(* PLC project conveyor_station.project, CODESYS CODESYS V3.5 SP22 Patch 4 *)
(* stored: creationDateTime 2026-11-23T00:04:54.4201515, modificationDateTime 2026-11-23T00:02:17.3371292 *)

PROGRAM PLC_PRG
  VAR
    START_BTN : BOOL;  (* physical NO button *)
    STOP_BTN : BOOL := TRUE;  (* physical NC button (TRUE = not pressed) *)
    RUN : BOOL;  (* memory bit: operator wants the conveyor running *)
    LAMP : BOOL;  (* warning lamp *)
    MOTOR : BOOL;  (* conveyor motor *)
    T1 : TON;  (* on-delay timer *)
    SENSOR : BOOL;  (* photo sensor: TRUE while a box blocks the beam *)
    RESET_BTN : BOOL;  (* operator resets the counter after swapping the crate *)
    C1 : CTU;  (* up-counter *)
    R1 : R_TRIG;  (* rising-edge detector for START *)
    START_EDGE : BOOL;  (* TRUE for one scan when START is pressed *)
    T2 : TON;  (* jam timer *)
    JAM : BOOL;  (* jam alarm (latched) *)
    ACK_BTN : BOOL;  (* operator acknowledges the alarm *)
  END_VAR

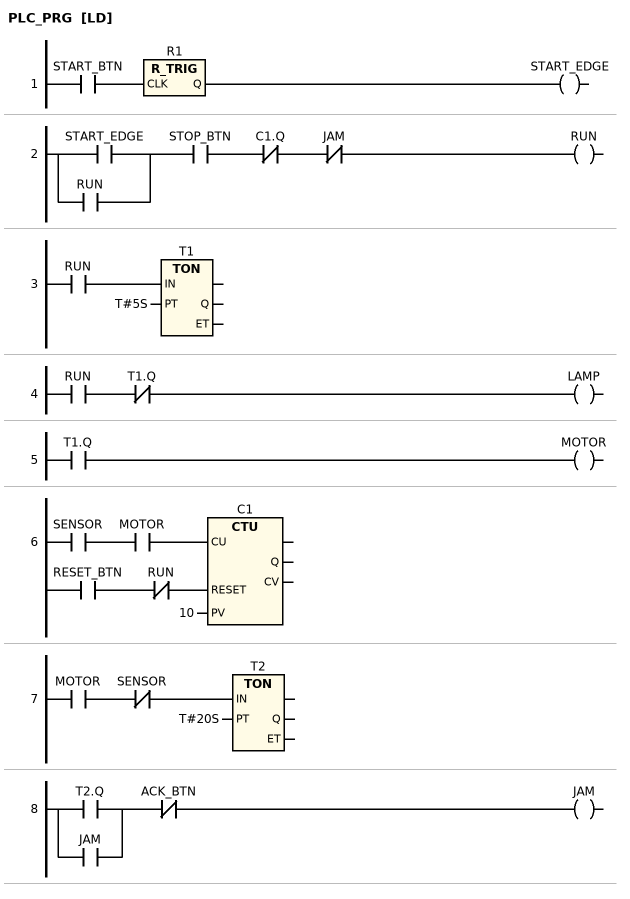
(* LD diagram, written out as Structured Text *)
(* --- network: Rising edge on START: prevents unexpected restart from a held/stuck button --- *)
R1(CLK := START_BTN);
START_EDGE := R1.Q;
(* --- network: Run latch: stopped by STOP, crate full (C1.Q) or jam (JAM) --- *)
RUN := (START_EDGE OR RUN) AND STOP_BTN AND NOT C1.Q AND NOT JAM;
(* --- network: 5 s warning timer before the conveyor moves --- *)
T1(IN := RUN, PT := T#5S);
(* --- network: Warning lamp ON during the 5 s countdown --- *)
LAMP := RUN AND NOT T1.Q;
(* --- network: Conveyor motor ON after the warning --- *)
MOTOR := T1.Q;
(* --- network: Box counter: counts only while the motor runs; crate full at 10; RESET only while stopped --- *)
C1(CU := SENSOR AND MOTOR, RESET := RESET_BTN AND NOT RUN, PV := 10);
(* --- network: Jam timer: motor running and no box at the sensor for 20 s --- *)
T2(IN := MOTOR AND NOT SENSOR, PT := T#20S);
(* --- network: Jam alarm latch: cleared only by ACK --- *)
JAM := (T2.Q OR JAM) AND NOT ACK_BTN;
END_PROGRAM
